Staubli VAL3: home.dtx

mdesc mNomSpeed
bool bEditAction
bool bEditIO
bool bEditTRAJ
bool bEditPROG
bool bEditFrame
bool bEditCycle
bool bEditSetting
bool bEditSpoint
bool bEditSzone
string sLib
num nLastStat
string sRobState
bool bExit
public string sVersion
bool bEditTcpTool
bool bLogMsg
